(* IEC 61131-3 sources: STAR-PLC-Agent/results/raw/six_task_fullflow_20261114/PUB007/generation/sim_00, 1 file *)

(* ---- test_program.st ---- *)
PROGRAM PLC_PRG
VAR
 BenchStep : UDINT := 0;
 BenchCalls : UDINT := 0;
 BenchDone : BOOL := FALSE;
 BenchUut0 : FB_Task;
 BenchUut1 : FB_Task;
 Binding_0_pumpGroup : ARRAY[1..5] OF ST_Pump;
 Binding_1_pumpGroup : ARRAY[1..5] OF ST_Pump;
 TraceIn_mode : ARRAY[0..7] OF BOOL;
 TraceIn_start : ARRAY[0..7] OF BOOL;
 TraceIn_stop : ARRAY[0..7] OF BOOL;
 TraceOut_pumpGroup_1_priority : ARRAY[0..7] OF INT;
 TraceOut_pumpGroup_1_selection : ARRAY[0..7] OF BOOL;
 TraceOut_pumpGroup_1_RunComd : ARRAY[0..7] OF BOOL;
 TraceOut_pumpGroup_2_priority : ARRAY[0..7] OF INT;
 TraceOut_pumpGroup_2_selection : ARRAY[0..7] OF BOOL;
 TraceOut_pumpGroup_2_RunComd : ARRAY[0..7] OF BOOL;
 TraceOut_pumpGroup_3_priority : ARRAY[0..7] OF INT;
 TraceOut_pumpGroup_3_selection : ARRAY[0..7] OF BOOL;
 TraceOut_pumpGroup_3_RunComd : ARRAY[0..7] OF BOOL;
 TraceOut_pumpGroup_4_priority : ARRAY[0..7] OF INT;
 TraceOut_pumpGroup_4_selection : ARRAY[0..7] OF BOOL;
 TraceOut_pumpGroup_4_RunComd : ARRAY[0..7] OF BOOL;
 TraceOut_pumpGroup_5_priority : ARRAY[0..7] OF INT;
 TraceOut_pumpGroup_5_selection : ARRAY[0..7] OF BOOL;
 TraceOut_pumpGroup_5_RunComd : ARRAY[0..7] OF BOOL;
END_VAR

IF NOT BenchDone THEN
 CASE BenchStep OF
 0:
   Binding_0_pumpGroup[1].priority := INT#1;
   Binding_0_pumpGroup[1].selection := TRUE;
   Binding_0_pumpGroup[1].RunComd := FALSE;
   Binding_0_pumpGroup[2].priority := INT#2;
   Binding_0_pumpGroup[2].selection := FALSE;
   Binding_0_pumpGroup[2].RunComd := FALSE;
   Binding_0_pumpGroup[3].priority := INT#3;
   Binding_0_pumpGroup[3].selection := TRUE;
   Binding_0_pumpGroup[3].RunComd := FALSE;
   Binding_0_pumpGroup[4].priority := INT#4;
   Binding_0_pumpGroup[4].selection := FALSE;
   Binding_0_pumpGroup[4].RunComd := FALSE;
   Binding_0_pumpGroup[5].priority := INT#5;
   Binding_0_pumpGroup[5].selection := FALSE;
   Binding_0_pumpGroup[5].RunComd := FALSE;
   BenchUut0.mode := FALSE;
   BenchUut0.start := TRUE;
   BenchUut0.stop := FALSE;
   TraceIn_mode[0] := BenchUut0.mode;
   TraceIn_start[0] := BenchUut0.start;
   TraceIn_stop[0] := BenchUut0.stop;
   BenchUut0(pumpGroup := Binding_0_pumpGroup);
   TraceOut_pumpGroup_1_priority[0] := Binding_0_pumpGroup[1].priority;
   TraceOut_pumpGroup_1_selection[0] := Binding_0_pumpGroup[1].selection;
   TraceOut_pumpGroup_1_RunComd[0] := Binding_0_pumpGroup[1].RunComd;
   TraceOut_pumpGroup_2_priority[0] := Binding_0_pumpGroup[2].priority;
   TraceOut_pumpGroup_2_selection[0] := Binding_0_pumpGroup[2].selection;
   TraceOut_pumpGroup_2_RunComd[0] := Binding_0_pumpGroup[2].RunComd;
   TraceOut_pumpGroup_3_priority[0] := Binding_0_pumpGroup[3].priority;
   TraceOut_pumpGroup_3_selection[0] := Binding_0_pumpGroup[3].selection;
   TraceOut_pumpGroup_3_RunComd[0] := Binding_0_pumpGroup[3].RunComd;
   TraceOut_pumpGroup_4_priority[0] := Binding_0_pumpGroup[4].priority;
   TraceOut_pumpGroup_4_selection[0] := Binding_0_pumpGroup[4].selection;
   TraceOut_pumpGroup_4_RunComd[0] := Binding_0_pumpGroup[4].RunComd;
   TraceOut_pumpGroup_5_priority[0] := Binding_0_pumpGroup[5].priority;
   TraceOut_pumpGroup_5_selection[0] := Binding_0_pumpGroup[5].selection;
   TraceOut_pumpGroup_5_RunComd[0] := Binding_0_pumpGroup[5].RunComd;
   BenchCalls := BenchCalls + 1;
 1:
   Binding_0_pumpGroup[1].priority := INT#1;
   Binding_0_pumpGroup[1].selection := FALSE;
   Binding_0_pumpGroup[1].RunComd := TRUE;
   Binding_0_pumpGroup[2].priority := INT#2;
   Binding_0_pumpGroup[2].selection := TRUE;
   Binding_0_pumpGroup[2].RunComd := FALSE;
   Binding_0_pumpGroup[3].priority := INT#3;
   Binding_0_pumpGroup[3].selection := FALSE;
   Binding_0_pumpGroup[3].RunComd := TRUE;
   Binding_0_pumpGroup[4].priority := INT#4;
   Binding_0_pumpGroup[4].selection := FALSE;
   Binding_0_pumpGroup[4].RunComd := FALSE;
   Binding_0_pumpGroup[5].priority := INT#5;
   Binding_0_pumpGroup[5].selection := FALSE;
   Binding_0_pumpGroup[5].RunComd := FALSE;
   BenchUut0.mode := FALSE;
   BenchUut0.start := FALSE;
   BenchUut0.stop := FALSE;
   TraceIn_mode[1] := BenchUut0.mode;
   TraceIn_start[1] := BenchUut0.start;
   TraceIn_stop[1] := BenchUut0.stop;
   BenchUut0(pumpGroup := Binding_0_pumpGroup);
   TraceOut_pumpGroup_1_priority[1] := Binding_0_pumpGroup[1].priority;
   TraceOut_pumpGroup_1_selection[1] := Binding_0_pumpGroup[1].selection;
   TraceOut_pumpGroup_1_RunComd[1] := Binding_0_pumpGroup[1].RunComd;
   TraceOut_pumpGroup_2_priority[1] := Binding_0_pumpGroup[2].priority;
   TraceOut_pumpGroup_2_selection[1] := Binding_0_pumpGroup[2].selection;
   TraceOut_pumpGroup_2_RunComd[1] := Binding_0_pumpGroup[2].RunComd;
   TraceOut_pumpGroup_3_priority[1] := Binding_0_pumpGroup[3].priority;
   TraceOut_pumpGroup_3_selection[1] := Binding_0_pumpGroup[3].selection;
   TraceOut_pumpGroup_3_RunComd[1] := Binding_0_pumpGroup[3].RunComd;
   TraceOut_pumpGroup_4_priority[1] := Binding_0_pumpGroup[4].priority;
   TraceOut_pumpGroup_4_selection[1] := Binding_0_pumpGroup[4].selection;
   TraceOut_pumpGroup_4_RunComd[1] := Binding_0_pumpGroup[4].RunComd;
   TraceOut_pumpGroup_5_priority[1] := Binding_0_pumpGroup[5].priority;
   TraceOut_pumpGroup_5_selection[1] := Binding_0_pumpGroup[5].selection;
   TraceOut_pumpGroup_5_RunComd[1] := Binding_0_pumpGroup[5].RunComd;
   BenchCalls := BenchCalls + 1;
 2:
   Binding_0_pumpGroup[1].priority := INT#1;
   Binding_0_pumpGroup[1].selection := FALSE;
   Binding_0_pumpGroup[1].RunComd := TRUE;
   Binding_0_pumpGroup[2].priority := INT#2;
   Binding_0_pumpGroup[2].selection := TRUE;
   Binding_0_pumpGroup[2].RunComd := FALSE;
   Binding_0_pumpGroup[3].priority := INT#3;
   Binding_0_pumpGroup[3].selection := FALSE;
   Binding_0_pumpGroup[3].RunComd := TRUE;
   Binding_0_pumpGroup[4].priority := INT#4;
   Binding_0_pumpGroup[4].selection := TRUE;
   Binding_0_pumpGroup[4].RunComd := FALSE;
   Binding_0_pumpGroup[5].priority := INT#5;
   Binding_0_pumpGroup[5].selection := FALSE;
   Binding_0_pumpGroup[5].RunComd := FALSE;
   BenchUut0.mode := FALSE;
   BenchUut0.start := TRUE;
   BenchUut0.stop := TRUE;
   TraceIn_mode[2] := BenchUut0.mode;
   TraceIn_start[2] := BenchUut0.start;
   TraceIn_stop[2] := BenchUut0.stop;
   BenchUut0(pumpGroup := Binding_0_pumpGroup);
   TraceOut_pumpGroup_1_priority[2] := Binding_0_pumpGroup[1].priority;
   TraceOut_pumpGroup_1_selection[2] := Binding_0_pumpGroup[1].selection;
   TraceOut_pumpGroup_1_RunComd[2] := Binding_0_pumpGroup[1].RunComd;
   TraceOut_pumpGroup_2_priority[2] := Binding_0_pumpGroup[2].priority;
   TraceOut_pumpGroup_2_selection[2] := Binding_0_pumpGroup[2].selection;
   TraceOut_pumpGroup_2_RunComd[2] := Binding_0_pumpGroup[2].RunComd;
   TraceOut_pumpGroup_3_priority[2] := Binding_0_pumpGroup[3].priority;
   TraceOut_pumpGroup_3_selection[2] := Binding_0_pumpGroup[3].selection;
   TraceOut_pumpGroup_3_RunComd[2] := Binding_0_pumpGroup[3].RunComd;
   TraceOut_pumpGroup_4_priority[2] := Binding_0_pumpGroup[4].priority;
   TraceOut_pumpGroup_4_selection[2] := Binding_0_pumpGroup[4].selection;
   TraceOut_pumpGroup_4_RunComd[2] := Binding_0_pumpGroup[4].RunComd;
   TraceOut_pumpGroup_5_priority[2] := Binding_0_pumpGroup[5].priority;
   TraceOut_pumpGroup_5_selection[2] := Binding_0_pumpGroup[5].selection;
   TraceOut_pumpGroup_5_RunComd[2] := Binding_0_pumpGroup[5].RunComd;
   BenchCalls := BenchCalls + 1;
 3:
   Binding_0_pumpGroup[1].priority := INT#1;
   Binding_0_pumpGroup[1].selection := FALSE;
   Binding_0_pumpGroup[1].RunComd := FALSE;
   Binding_0_pumpGroup[2].priority := INT#2;
   Binding_0_pumpGroup[2].selection := FALSE;
   Binding_0_pumpGroup[2].RunComd := FALSE;
   Binding_0_pumpGroup[3].priority := INT#3;
   Binding_0_pumpGroup[3].selection := FALSE;
   Binding_0_pumpGroup[3].RunComd := FALSE;
   Binding_0_pumpGroup[4].priority := INT#4;
   Binding_0_pumpGroup[4].selection := FALSE;
   Binding_0_pumpGroup[4].RunComd := FALSE;
   Binding_0_pumpGroup[5].priority := INT#5;
   Binding_0_pumpGroup[5].selection := TRUE;
   Binding_0_pumpGroup[5].RunComd := FALSE;
   BenchUut0.mode := FALSE;
   BenchUut0.start := TRUE;
   BenchUut0.stop := FALSE;
   TraceIn_mode[3] := BenchUut0.mode;
   TraceIn_start[3] := BenchUut0.start;
   TraceIn_stop[3] := BenchUut0.stop;
   BenchUut0(pumpGroup := Binding_0_pumpGroup);
   TraceOut_pumpGroup_1_priority[3] := Binding_0_pumpGroup[1].priority;
   TraceOut_pumpGroup_1_selection[3] := Binding_0_pumpGroup[1].selection;
   TraceOut_pumpGroup_1_RunComd[3] := Binding_0_pumpGroup[1].RunComd;
   TraceOut_pumpGroup_2_priority[3] := Binding_0_pumpGroup[2].priority;
   TraceOut_pumpGroup_2_selection[3] := Binding_0_pumpGroup[2].selection;
   TraceOut_pumpGroup_2_RunComd[3] := Binding_0_pumpGroup[2].RunComd;
   TraceOut_pumpGroup_3_priority[3] := Binding_0_pumpGroup[3].priority;
   TraceOut_pumpGroup_3_selection[3] := Binding_0_pumpGroup[3].selection;
   TraceOut_pumpGroup_3_RunComd[3] := Binding_0_pumpGroup[3].RunComd;
   TraceOut_pumpGroup_4_priority[3] := Binding_0_pumpGroup[4].priority;
   TraceOut_pumpGroup_4_selection[3] := Binding_0_pumpGroup[4].selection;
   TraceOut_pumpGroup_4_RunComd[3] := Binding_0_pumpGroup[4].RunComd;
   TraceOut_pumpGroup_5_priority[3] := Binding_0_pumpGroup[5].priority;
   TraceOut_pumpGroup_5_selection[3] := Binding_0_pumpGroup[5].selection;
   TraceOut_pumpGroup_5_RunComd[3] := Binding_0_pumpGroup[5].RunComd;
   BenchCalls := BenchCalls + 1;
 4:
   Binding_1_pumpGroup[1].priority := INT#10;
   Binding_1_pumpGroup[1].selection := TRUE;
   Binding_1_pumpGroup[1].RunComd := FALSE;
   Binding_1_pumpGroup[2].priority := INT#20;
   Binding_1_pumpGroup[2].selection := FALSE;
   Binding_1_pumpGroup[2].RunComd := FALSE;
   Binding_1_pumpGroup[3].priority := INT#20;
   Binding_1_pumpGroup[3].selection := FALSE;
   Binding_1_pumpGroup[3].RunComd := FALSE;
   Binding_1_pumpGroup[4].priority := INT#20;
   Binding_1_pumpGroup[4].selection := TRUE;
   Binding_1_pumpGroup[4].RunComd := FALSE;
   Binding_1_pumpGroup[5].priority := INT#30;
   Binding_1_pumpGroup[5].selection := FALSE;
   Binding_1_pumpGroup[5].RunComd := FALSE;
   BenchUut1.mode := TRUE;
   BenchUut1.start := TRUE;
   BenchUut1.stop := FALSE;
   TraceIn_mode[4] := BenchUut1.mode;
   TraceIn_start[4] := BenchUut1.start;
   TraceIn_stop[4] := BenchUut1.stop;
   BenchUut1(pumpGroup := Binding_1_pumpGroup);
   TraceOut_pumpGroup_1_priority[4] := Binding_1_pumpGroup[1].priority;
   TraceOut_pumpGroup_1_selection[4] := Binding_1_pumpGroup[1].selection;
   TraceOut_pumpGroup_1_RunComd[4] := Binding_1_pumpGroup[1].RunComd;
   TraceOut_pumpGroup_2_priority[4] := Binding_1_pumpGroup[2].priority;
   TraceOut_pumpGroup_2_selection[4] := Binding_1_pumpGroup[2].selection;
   TraceOut_pumpGroup_2_RunComd[4] := Binding_1_pumpGroup[2].RunComd;
   TraceOut_pumpGroup_3_priority[4] := Binding_1_pumpGroup[3].priority;
   TraceOut_pumpGroup_3_selection[4] := Binding_1_pumpGroup[3].selection;
   TraceOut_pumpGroup_3_RunComd[4] := Binding_1_pumpGroup[3].RunComd;
   TraceOut_pumpGroup_4_priority[4] := Binding_1_pumpGroup[4].priority;
   TraceOut_pumpGroup_4_selection[4] := Binding_1_pumpGroup[4].selection;
   TraceOut_pumpGroup_4_RunComd[4] := Binding_1_pumpGroup[4].RunComd;
   TraceOut_pumpGroup_5_priority[4] := Binding_1_pumpGroup[5].priority;
   TraceOut_pumpGroup_5_selection[4] := Binding_1_pumpGroup[5].selection;
   TraceOut_pumpGroup_5_RunComd[4] := Binding_1_pumpGroup[5].RunComd;
   BenchCalls := BenchCalls + 1;
 5:
   Binding_1_pumpGroup[1].priority := INT#50;
   Binding_1_pumpGroup[1].selection := FALSE;
   Binding_1_pumpGroup[1].RunComd := FALSE;
   Binding_1_pumpGroup[2].priority := INT#1;
   Binding_1_pumpGroup[2].selection := TRUE;
   Binding_1_pumpGroup[2].RunComd := TRUE;
   Binding_1_pumpGroup[3].priority := INT#1;
   Binding_1_pumpGroup[3].selection := FALSE;
   Binding_1_pumpGroup[3].RunComd := TRUE;
   Binding_1_pumpGroup[4].priority := INT#1;
   Binding_1_pumpGroup[4].selection := FALSE;
   Binding_1_pumpGroup[4].RunComd := FALSE;
   Binding_1_pumpGroup[5].priority := INT#1;
   Binding_1_pumpGroup[5].selection := FALSE;
   Binding_1_pumpGroup[5].RunComd := TRUE;
   BenchUut1.mode := TRUE;
   BenchUut1.start := FALSE;
   BenchUut1.stop := FALSE;
   TraceIn_mode[5] := BenchUut1.mode;
   TraceIn_start[5] := BenchUut1.start;
   TraceIn_stop[5] := BenchUut1.stop;
   BenchUut1(pumpGroup := Binding_1_pumpGroup);
   TraceOut_pumpGroup_1_priority[5] := Binding_1_pumpGroup[1].priority;
   TraceOut_pumpGroup_1_selection[5] := Binding_1_pumpGroup[1].selection;
   TraceOut_pumpGroup_1_RunComd[5] := Binding_1_pumpGroup[1].RunComd;
   TraceOut_pumpGroup_2_priority[5] := Binding_1_pumpGroup[2].priority;
   TraceOut_pumpGroup_2_selection[5] := Binding_1_pumpGroup[2].selection;
   TraceOut_pumpGroup_2_RunComd[5] := Binding_1_pumpGroup[2].RunComd;
   TraceOut_pumpGroup_3_priority[5] := Binding_1_pumpGroup[3].priority;
   TraceOut_pumpGroup_3_selection[5] := Binding_1_pumpGroup[3].selection;
   TraceOut_pumpGroup_3_RunComd[5] := Binding_1_pumpGroup[3].RunComd;
   TraceOut_pumpGroup_4_priority[5] := Binding_1_pumpGroup[4].priority;
   TraceOut_pumpGroup_4_selection[5] := Binding_1_pumpGroup[4].selection;
   TraceOut_pumpGroup_4_RunComd[5] := Binding_1_pumpGroup[4].RunComd;
   TraceOut_pumpGroup_5_priority[5] := Binding_1_pumpGroup[5].priority;
   TraceOut_pumpGroup_5_selection[5] := Binding_1_pumpGroup[5].selection;
   TraceOut_pumpGroup_5_RunComd[5] := Binding_1_pumpGroup[5].RunComd;
   BenchCalls := BenchCalls + 1;
 6:
   Binding_1_pumpGroup[1].priority := INT#50;
   Binding_1_pumpGroup[1].selection := FALSE;
   Binding_1_pumpGroup[1].RunComd := FALSE;
   Binding_1_pumpGroup[2].priority := INT#1;
   Binding_1_pumpGroup[2].selection := TRUE;
   Binding_1_pumpGroup[2].RunComd := TRUE;
   Binding_1_pumpGroup[3].priority := INT#1;
   Binding_1_pumpGroup[3].selection := FALSE;
   Binding_1_pumpGroup[3].RunComd := TRUE;
   Binding_1_pumpGroup[4].priority := INT#1;
   Binding_1_pumpGroup[4].selection := FALSE;
   Binding_1_pumpGroup[4].RunComd := FALSE;
   Binding_1_pumpGroup[5].priority := INT#1;
   Binding_1_pumpGroup[5].selection := FALSE;
   Binding_1_pumpGroup[5].RunComd := TRUE;
   BenchUut1.mode := TRUE;
   BenchUut1.start := TRUE;
   BenchUut1.stop := FALSE;
   TraceIn_mode[6] := BenchUut1.mode;
   TraceIn_start[6] := BenchUut1.start;
   TraceIn_stop[6] := BenchUut1.stop;
   BenchUut1(pumpGroup := Binding_1_pumpGroup);
   TraceOut_pumpGroup_1_priority[6] := Binding_1_pumpGroup[1].priority;
   TraceOut_pumpGroup_1_selection[6] := Binding_1_pumpGroup[1].selection;
   TraceOut_pumpGroup_1_RunComd[6] := Binding_1_pumpGroup[1].RunComd;
   TraceOut_pumpGroup_2_priority[6] := Binding_1_pumpGroup[2].priority;
   TraceOut_pumpGroup_2_selection[6] := Binding_1_pumpGroup[2].selection;
   TraceOut_pumpGroup_2_RunComd[6] := Binding_1_pumpGroup[2].RunComd;
   TraceOut_pumpGroup_3_priority[6] := Binding_1_pumpGroup[3].priority;
   TraceOut_pumpGroup_3_selection[6] := Binding_1_pumpGroup[3].selection;
   TraceOut_pumpGroup_3_RunComd[6] := Binding_1_pumpGroup[3].RunComd;
   TraceOut_pumpGroup_4_priority[6] := Binding_1_pumpGroup[4].priority;
   TraceOut_pumpGroup_4_selection[6] := Binding_1_pumpGroup[4].selection;
   TraceOut_pumpGroup_4_RunComd[6] := Binding_1_pumpGroup[4].RunComd;
   TraceOut_pumpGroup_5_priority[6] := Binding_1_pumpGroup[5].priority;
   TraceOut_pumpGroup_5_selection[6] := Binding_1_pumpGroup[5].selection;
   TraceOut_pumpGroup_5_RunComd[6] := Binding_1_pumpGroup[5].RunComd;
   BenchCalls := BenchCalls + 1;
 7:
   Binding_1_pumpGroup[1].priority := INT#50;
   Binding_1_pumpGroup[1].selection := FALSE;
   Binding_1_pumpGroup[1].RunComd := TRUE;
   Binding_1_pumpGroup[2].priority := INT#1;
   Binding_1_pumpGroup[2].selection := TRUE;
   Binding_1_pumpGroup[2].RunComd := TRUE;
   Binding_1_pumpGroup[3].priority := INT#1;
   Binding_1_pumpGroup[3].selection := FALSE;
   Binding_1_pumpGroup[3].RunComd := TRUE;
   Binding_1_pumpGroup[4].priority := INT#1;
   Binding_1_pumpGroup[4].selection := FALSE;
   Binding_1_pumpGroup[4].RunComd := FALSE;
   Binding_1_pumpGroup[5].priority := INT#1;
   Binding_1_pumpGroup[5].selection := FALSE;
   Binding_1_pumpGroup[5].RunComd := FALSE;
   BenchUut1.mode := TRUE;
   BenchUut1.start := TRUE;
   BenchUut1.stop := TRUE;
   TraceIn_mode[7] := BenchUut1.mode;
   TraceIn_start[7] := BenchUut1.start;
   TraceIn_stop[7] := BenchUut1.stop;
   BenchUut1(pumpGroup := Binding_1_pumpGroup);
   TraceOut_pumpGroup_1_priority[7] := Binding_1_pumpGroup[1].priority;
   TraceOut_pumpGroup_1_selection[7] := Binding_1_pumpGroup[1].selection;
   TraceOut_pumpGroup_1_RunComd[7] := Binding_1_pumpGroup[1].RunComd;
   TraceOut_pumpGroup_2_priority[7] := Binding_1_pumpGroup[2].priority;
   TraceOut_pumpGroup_2_selection[7] := Binding_1_pumpGroup[2].selection;
   TraceOut_pumpGroup_2_RunComd[7] := Binding_1_pumpGroup[2].RunComd;
   TraceOut_pumpGroup_3_priority[7] := Binding_1_pumpGroup[3].priority;
   TraceOut_pumpGroup_3_selection[7] := Binding_1_pumpGroup[3].selection;
   TraceOut_pumpGroup_3_RunComd[7] := Binding_1_pumpGroup[3].RunComd;
   TraceOut_pumpGroup_4_priority[7] := Binding_1_pumpGroup[4].priority;
   TraceOut_pumpGroup_4_selection[7] := Binding_1_pumpGroup[4].selection;
   TraceOut_pumpGroup_4_RunComd[7] := Binding_1_pumpGroup[4].RunComd;
   TraceOut_pumpGroup_5_priority[7] := Binding_1_pumpGroup[5].priority;
   TraceOut_pumpGroup_5_selection[7] := Binding_1_pumpGroup[5].selection;
   TraceOut_pumpGroup_5_RunComd[7] := Binding_1_pumpGroup[5].RunComd;
   BenchCalls := BenchCalls + 1;
 END_CASE;
 BenchStep := BenchStep + 1;
 IF BenchStep >= 8 THEN BenchDone := TRUE; END_IF;
END_IF;
END_PROGRAM
